// TIA Portal V14 SP1 export
// export: Created 2000-01-01T00:00:00.0000000Z, ExportSetting None
DATA_BLOCK "MCP_RC_DB4"   // DB9804
{ S7_Optimized_Access := 'TRUE' }
   VAR
      "A" : "MCP_RC_UDT2";
      "B" : "MCP_RC_UDT2";
   END_VAR
BEGIN
END_DATA_BLOCK
